(* IEC 61131-3 sources: Codesys_IAP/Demo/PLC1/PLC 1 Simulatie Ladder StructuredTekst IOStructures 2V0_tekst/Programma Structured Text/UitvoerGootClass, 9 files *)

(* ---- cycle.st ---- *)
(*#### DECLARATIE ####*)
// Datum : 17 december 2020, Auteur: Gerard Harkema
METHOD cycle
VAR_INPUT
END_VAR

(*#### IMPLEMENTATIE ####*)
CASE eState OF
//	uitvoerGootStates.idle:
//	uitvoerGootStates.is_in:
	uitvoerGootStates.ga_in:
	IF IO.Ix_UitvoerGootIsIn THEN
		eState := uitvoerGootStates.is_in;
	END_IF

//	uitvoerGootStates.is_uit:
	uitvoerGootStates.ga_uit:
	IF IO.Ix_UitvoerGootIsUit THEN
		eState := uitvoerGootStates.is_uit;
	END_IF
//	uitvoerGootStates.error:
END_CASE

(* ---- gaIn.st ---- *)
(*#### DECLARATIE ####*)
// Datum : 17 december 2020, Auteur: Gerard Harkema
METHOD gaIn
VAR_INPUT
END_VAR

(*#### IMPLEMENTATIE ####*)
IF NOT (eState = uitvoerGootStates.is_uit) THEN
	eState := uitvoerGootStates.error;
	return;
END_IF

IO.Qx_UitvoerGootUit := FALSE;
eState := uitvoerGootStates.ga_in;

(* ---- gaUit.st ---- *)
(*#### DECLARATIE ####*)
// Datum : 17 december 2020, Auteur: Gerard Harkema
METHOD gaUit
VAR_INPUT
END_VAR

(*#### IMPLEMENTATIE ####*)
IF NOT (eState = uitvoerGootStates.is_in) THEN
	eState := uitvoerGootStates.error;
	return;
END_IF

IO.Qx_UitvoerGootUit := TRUE;
eState := uitvoerGootStates.ga_uit;

(* ---- initialize.st ---- *)
(*#### DECLARATIE ####*)
// Datum : 17 december 2020, Auteur: Gerard Harkema
METHOD initialize
VAR_INPUT
	IORef			: REFERENCE TO uitvoerGootIO;

END_VAR

(*#### IMPLEMENTATIE ####*)
//Pusher uitvoergoot is in
IO 	REF=	IORef;
eState := uitvoerGootStates.ga_in;

(* ---- isError.st ---- *)
(*#### DECLARATIE ####*)
// Datum : 17 december 2020, Auteur: Gerard Harkema
METHOD isError : BOOL
VAR_INPUT
END_VAR

(*#### IMPLEMENTATIE ####*)
isError := (eState = uitvoerGootStates.error);

(* ---- isIn.st ---- *)
(*#### DECLARATIE ####*)
// Datum : 17 december 2020, Auteur: Gerard Harkema
METHOD isIn : BOOL
VAR_INPUT
END_VAR

(*#### IMPLEMENTATIE ####*)
isIn := (eState = uitvoerGootStates.is_in);

(* ---- isUit.st ---- *)
(*#### DECLARATIE ####*)
// Datum : 17 december 2020, Auteur: Gerard Harkema
METHOD isUit : BOOL
VAR_INPUT
END_VAR

(*#### IMPLEMENTATIE ####*)
isUit := (eState = uitvoerGootStates.is_uit);

(* ---- noodstop.st ---- *)
(*#### DECLARATIE ####*)
// Datum : 17 december 2020, Auteur: Gerard Harkema
METHOD noodstop
VAR_INPUT
END_VAR

(*#### IMPLEMENTATIE ####*)
IO.Qx_UitvoerGootUit := FALSE;
eState := uitvoerGootStates.error;

(* ---- reset.st ---- *)
(*#### DECLARATIE ####*)
// Datum : 17 december 2020, Auteur: Gerard Harkema
METHOD reset
VAR_INPUT
END_VAR

(*#### IMPLEMENTATIE ####*)
IO.Qx_UitvoerGootUit := FALSE;
eState := uitvoerGootStates.ga_in;
